// TIA Portal V21 export
GraphicList "GL_Bit"  ListRange=Bit
  GraphicListEntry   EntryType=SingleValue, Picture=G_EMF
  GraphicListEntry   EntryType=SingleValue, From=1, To=1, Picture=G_WMF
